Fanuc KAREL source: kt00574.KL

-- PROVISIONAL review KL for V1013-1; original PC SHA256 785f66c838c69f222c2c88783ebe3c42a72abb40eabff482d01a5788188dc16e
-- Incomplete behavior may be omitted. Consult companion uncertainty JSON. Do not deploy.
PROGRAM KT00574
%NOLOCKGROUP
VAR
  R1 : REAL
-- UNRESOLVED_DECL V2 type=000013
-- UNRESOLVED_DECL OUT type=000013
BEGIN
  -- UNRESOLVED_PC offsets 5-16; opcodes 2E,23
  -- UNRESOLVED_PC offsets 21-36; opcodes 2E,22,32,35
  -- UNRESOLVED_PC offsets 41-63; opcodes 21,49,90,4A
  -- UNRESOLVED_PC offsets 68-72; opcodes 7F
END KT00574
